Staubli VAL3: areaCheck.pgx

public program areaCheck()
  local num l_i
begin
  for l_i = 0 to size(safeData:zZoneItem)-1
    if safeData:zZoneItem[l_i].bActive
      call computeArea(l_i)
    endIf
  endFor

end
